(* IEC 61131-3 sources: PortalRobot/Portal_robot/Device/application/FB, 43 files *)

(* ---- F_GEOMETRY_EVENT.st ---- *)
FUNCTION F_GEOMETRY_EVENT : BOOL
VAR_INPUT
	Call : ST_GEOMETRY_CALL;
END_VAR
VAR
	uiIndex : UINT;
END_VAR

// --- BEGIN IMPLEMENTATION ---

// Один PLC-скан, единый владелец номера. Поля записываются раньше Seq.
Persistent_Value.udiEventSequence := Persistent_Value.udiEventSequence + UDINT#1;
IF Persistent_Value.udiEventSequence = UDINT#0 THEN Persistent_Value.udiEventSequence := UDINT#1; END_IF;
uiIndex := UDINT_TO_UINT((Persistent_Value.udiEventSequence - UDINT#1) MOD UDINT#100) + UINT#1;
GVL_GEOMETRY_CONTROL.astEvents[uiIndex].udiSequence := UDINT#0;
GVL_GEOMETRY_CONTROL.astEvents[uiIndex].Call := Call;
GVL_GEOMETRY_CONTROL.astEvents[uiIndex].udiTimeMs := GVL_HMI.udiHmiCommandClockMs;
GVL_GEOMETRY_CONTROL.astEvents[uiIndex].uiEnvironment := GVL_GEOMETRY_CONTROL.uiEnvironment;
GVL_GEOMETRY_CONTROL.astEvents[uiIndex].udiSequence := Persistent_Value.udiEventSequence;
F_GEOMETRY_EVENT := TRUE;

(* ---- F_GEOMETRY_SELECT_STATION.st ---- *)
FUNCTION F_GEOMETRY_SELECT_STATION : UINT
VAR_INPUT
	xRequireFree : BOOL;
	uiMachine : UINT := UINT#0; // Станок-источник; 0 — общая проверка доступности
END_VAR
VAR
	uiTry : UINT;
	uiStation : UINT;
END_VAR

// --- BEGIN IMPLEMENTATION ---

F_GEOMETRY_SELECT_STATION := UINT#0;
// С1/С2 предпочитают ГК1, С3 — ГК2. История доставок и магазины не участвуют.
uiStation := UINT#1;
IF uiMachine = UINT#3 THEN uiStation := UINT#2; END_IF;
FOR uiTry := UINT#1 TO UINT#2 DO
	// Вторым проверяем другой ГК, если предпочтительный не прошёл допуск.
	IF uiTry = UINT#2 THEN uiStation := UINT#3 - uiStation; END_IF;
	IF (F_GEOMETRY_SELECT_STATION = UINT#0) AND GVL_GEOMETRY_CONTROL.xSupported
	AND GVL_GEOMETRY_CONTROL.astStatus[uiStation].xEnabled
	AND NOT GVL_GEOMETRY_CONTROL.astStatus[uiStation].xDisablePending
	AND GVL_GEOMETRY_CONTROL.astStatus[uiStation].xConfigured
	AND NOT GVL_GEOMETRY_CONTROL.astStatus[uiStation].xError
	AND (GVL_GEOMETRY_CONTROL.astStatus[uiStation].uiState <> UINT#5) THEN
		IF NOT xRequireFree OR GVL_GEOMETRY_CONTROL.astStatus[uiStation].xReady THEN F_GEOMETRY_SELECT_STATION := uiStation; END_IF;
	END_IF;
END_FOR;

(* ---- F_GEOMETRY_TAKE_DETAIL.st ---- *)
FUNCTION F_GEOMETRY_TAKE_DETAIL : BOOL
VAR_INPUT
	uiMachine : UINT;
	uiProductType : UINT;
END_VAR
VAR
	Call : ST_GEOMETRY_CALL;
	EmptyCall : ST_GEOMETRY_CALL;
END_VAR

// --- BEGIN IMPLEMENTATION ---

F_GEOMETRY_TAKE_DETAIL := FALSE;
IF (uiMachine >= UINT#1) AND (uiMachine <= UINT#3) THEN
	// Считаем подтверждённую выгрузку ровно один раз, а не уровень Ready каждый скан.
	// Ожидающая выборка сохраняет счётчик до фактического взятия своей детали.
	IF (GVL_GEOMETRY_CONTROL.astCalls[uiMachine].uiState <> UINT#1)
	AND GVL_GEOMETRY_CONTROL.xSupported AND Persistent_Value.xAutoEnabled
	AND (GVL_GEOMETRY_CONTROL.astStatus[1].xEnabled OR GVL_GEOMETRY_CONTROL.astStatus[2].xEnabled) THEN
		GVL_GEOMETRY_CONTROL.auiActiveCount[uiMachine] := MIN(UINT#10000, GVL_GEOMETRY_CONTROL.auiActiveCount[uiMachine] + UINT#1);
		IF GVL_GEOMETRY_CONTROL.auiActiveCount[uiMachine] >= Persistent_Value.auiPeriod[uiMachine] THEN
			IF (GVL_GEOMETRY_CONTROL.astCalls[uiMachine].uiState <> UINT#2)
			AND (GVL_GEOMETRY_CONTROL.astCalls[uiMachine].uiState <> UINT#3) THEN
				Persistent_Value.udiNextCallId := Persistent_Value.udiNextCallId + UDINT#1;
				IF Persistent_Value.udiNextCallId = UDINT#0 THEN Persistent_Value.udiNextCallId := UDINT#1; END_IF;
				Call := EmptyCall; Call.udiId := Persistent_Value.udiNextCallId;
				Call.uiMachine := uiMachine; Call.uiProductType := uiProductType; Call.uiState := UINT#1;
				GVL_GEOMETRY_CONTROL.astCalls[uiMachine] := Call; F_GEOMETRY_EVENT(Call := Call);
			ELSE
				GVL_GEOMETRY_CONTROL.auiActiveCount[uiMachine] := UINT#0;
			END_IF;
		END_IF;
	END_IF;
	// Подхватываем вызов обслуживаемого станка независимо от вызовов других станков.
	// Повторная проверка после выезда также допускает поздний вызов своей детали.
	IF GVL_GEOMETRY_CONTROL.astCalls[uiMachine].uiState = UINT#1 THEN
		GVL_GEOMETRY_CONTROL.auiActiveCount[uiMachine] := UINT#0;
		GVL_GEOMETRY_CONTROL.astCalls[uiMachine].uiProductType := uiProductType;
		GVL_GEOMETRY_CONTROL.astCalls[uiMachine].uiState := UINT#2;
		F_GEOMETRY_EVENT(Call := GVL_GEOMETRY_CONTROL.astCalls[uiMachine]);
		F_GEOMETRY_TAKE_DETAIL := TRUE;
	END_IF;
END_IF;

(* ---- F_MAGAZINE_FRAME.st ---- *)
FUNCTION F_MAGAZINE_FRAME : ST_MAGAZINE_FRAME
VAR_INPUT
	stOrigin : ST_POINT;
	stCalibration : ST_MAGAZINE_CALIBRATION;
	uiRows : UINT;
	uiColumns : UINT;
	lrPitchX : LREAL;
	lrPitchY : LREAL;
END_VAR
VAR
	stFrame : ST_MAGAZINE_FRAME;
	stVectorAB : ST_MAGAZINE_VECTOR;
	stVectorAC : ST_MAGAZINE_VECTOR;
	stPlaneNormal : ST_MAGAZINE_VECTOR;
	lrVectorABLength : LREAL;
	lrPlaneNormalLength : LREAL;
END_VAR

// --- BEGIN IMPLEMENTATION ---

// Одноточечный режим сохраняет прежние направления мировых X/Y.
stFrame.stAxisX.X := 1.0; stFrame.stAxisX.Y := 0.0; stFrame.stAxisX.Z := 0.0;
stFrame.stAxisY.X := 0.0; stFrame.stAxisY.Y := 1.0; stFrame.stAxisY.Z := 0.0;
stFrame.stAxisZ.X := 0.0; stFrame.stAxisZ.Y := 0.0; stFrame.stAxisZ.Z := 1.0;
stFrame.xReady := FALSE;
stFrame.uiReason := UINT#0;
IF NOT stOrigin.xConfigured
OR (stOrigin.MagazineSafeZ = 0.0) OR (stOrigin.MagazineChangeZ = 0.0) THEN
	stFrame.uiReason := UINT#1;
ELSIF ((stCalibration.uiMethod <> UINT#1) AND (stCalibration.uiMethod <> UINT#3))
OR (uiRows = UINT#0) OR (uiColumns = UINT#0)
OR NOT ((lrPitchX >= 1.0) AND (lrPitchX <= 5000.0)
	AND (lrPitchY >= 1.0) AND (lrPitchY <= 5000.0)) THEN
	stFrame.uiReason := UINT#2;
ELSIF stCalibration.uiMethod = UINT#1 THEN
	stFrame.xReady := TRUE;
ELSIF (uiRows < UINT#2) OR (uiColumns < UINT#2) THEN
	stFrame.uiReason := UINT#2;
ELSIF NOT stCalibration.astReference[1].xConfigured
OR NOT stCalibration.astReference[2].xConfigured THEN
	stFrame.uiReason := UINT#3;
ELSE
	stVectorAB.X := stCalibration.astReference[1].X - stOrigin.X;
	stVectorAB.Y := stCalibration.astReference[1].Y - stOrigin.Y;
	stVectorAB.Z := stCalibration.astReference[1].Z - stOrigin.Z;
	stVectorAC.X := stCalibration.astReference[2].X - stOrigin.X;
	stVectorAC.Y := stCalibration.astReference[2].Y - stOrigin.Y;
	stVectorAC.Z := stCalibration.astReference[2].Z - stOrigin.Z;
	stPlaneNormal.X := stVectorAB.Y * stVectorAC.Z - stVectorAB.Z * stVectorAC.Y;
	stPlaneNormal.Y := stVectorAB.Z * stVectorAC.X - stVectorAB.X * stVectorAC.Z;
	stPlaneNormal.Z := stVectorAB.X * stVectorAC.Y - stVectorAB.Y * stVectorAC.X;
	lrVectorABLength := SQRT(stVectorAB.X * stVectorAB.X + stVectorAB.Y * stVectorAB.Y + stVectorAB.Z * stVectorAB.Z);
	lrPlaneNormalLength := SQRT(stPlaneNormal.X * stPlaneNormal.X + stPlaneNormal.Y * stPlaneNormal.Y + stPlaneNormal.Z * stPlaneNormal.Z);
	// Только математическая определённость: допуски размеров/углов не применяются.
	IF (lrVectorABLength > 0.0) AND (lrPlaneNormalLength > 0.0) THEN
		stFrame.stAxisX.X := stVectorAB.X / lrVectorABLength;
		stFrame.stAxisX.Y := stVectorAB.Y / lrVectorABLength;
		stFrame.stAxisX.Z := stVectorAB.Z / lrVectorABLength;
		stFrame.stAxisZ.X := stPlaneNormal.X / lrPlaneNormalLength;
		stFrame.stAxisZ.Y := stPlaneNormal.Y / lrPlaneNormalLength;
		stFrame.stAxisZ.Z := stPlaneNormal.Z / lrPlaneNormalLength;
		stFrame.stAxisY.X := stFrame.stAxisZ.Y * stFrame.stAxisX.Z - stFrame.stAxisZ.Z * stFrame.stAxisX.Y;
		stFrame.stAxisY.Y := stFrame.stAxisZ.Z * stFrame.stAxisX.X - stFrame.stAxisZ.X * stFrame.stAxisX.Z;
		stFrame.stAxisY.Z := stFrame.stAxisZ.X * stFrame.stAxisX.Y - stFrame.stAxisZ.Y * stFrame.stAxisX.X;
		// Сравнения также не принимают NaN/Inf после нечисловых входных данных.
		stFrame.xReady := (ABS(stFrame.stAxisX.X) <= 2.0) AND (ABS(stFrame.stAxisX.Y) <= 2.0)
			AND (ABS(stFrame.stAxisX.Z) <= 2.0) AND (ABS(stFrame.stAxisY.X) <= 2.0)
			AND (ABS(stFrame.stAxisY.Y) <= 2.0) AND (ABS(stFrame.stAxisY.Z) <= 2.0)
			AND (ABS(stFrame.stAxisZ.X) <= 2.0) AND (ABS(stFrame.stAxisZ.Y) <= 2.0)
			AND (ABS(stFrame.stAxisZ.Z) <= 2.0)
			AND ((stFrame.stAxisX.X * stFrame.stAxisX.X + stFrame.stAxisX.Y * stFrame.stAxisX.Y + stFrame.stAxisX.Z * stFrame.stAxisX.Z) > 0.0)
			AND ((stFrame.stAxisZ.X * stFrame.stAxisZ.X + stFrame.stAxisZ.Y * stFrame.stAxisZ.Y + stFrame.stAxisZ.Z * stFrame.stAxisZ.Z) > 0.0);
	END_IF;
	IF NOT stFrame.xReady THEN stFrame.uiReason := UINT#4; END_IF;
END_IF;
F_MAGAZINE_FRAME := stFrame;

(* ---- FB_ALARM_HORN.st ---- *)
FUNCTION_BLOCK FB_ALARM_HORN
VAR_INPUT
    astSource : ARRAY [1..22] OF ST_ALARM_SOURCE_DATA;
    tDuration : TIME := T#2S;
END_VAR
VAR_OUTPUT
    xSound : BOOL;
END_VAR
VAR
    adwPrevious : ARRAY [1..22] OF DWORD;
    uiSource : UINT;
    xNewAlarm : BOOL;
    xActive : BOOL;
    tLatchedDuration : TIME;
    tonSound : TON;
END_VAR

// --- BEGIN IMPLEMENTATION ---

// Предупреждения не входят в dwAlarmActive. Новая авария другого источника/бита
// тоже запускает звук, даже когда общая xAlarmActive уже была TRUE.
xNewAlarm := FALSE;
FOR uiSource := 1 TO 22 DO
    IF (astSource[uiSource].dwAlarmActive AND NOT adwPrevious[uiSource]) <> DWORD#0 THEN
        xNewAlarm := TRUE;
    END_IF;
    adwPrevious[uiSource] := astSource[uiSource].dwAlarmActive;
END_FOR;
IF tDuration <= T#0MS THEN
    xActive := FALSE;
ELSIF xNewAlarm THEN
    xActive := TRUE;
    tLatchedDuration := tDuration;
    // Сброс и запуск TON в этом же скане: новая авария начинает полный интервал.
    tonSound(IN := FALSE, PT := tLatchedDuration);
END_IF;
tonSound(IN := xActive, PT := tLatchedDuration);
IF tonSound.Q THEN
    xActive := FALSE;
END_IF;
xSound := xActive;

(* ---- FB_ALARM_MANAGER.st ---- *)
FUNCTION_BLOCK FB_ALARM_MANAGER
VAR_INPUT
	xResetWarnings : BOOL; // Сброс накопленных предупреждений
    xControllerWarningResetAllowed : BOOL; // 5C нельзя подтвердить до исчезновения свежей причины.
	astAdditionalCellWarning : ARRAY [1..2] OF ST_WARNING_EVENT; // Конфигуратор и ГК: независимые события источника CELL
END_VAR
VAR_IN_OUT
	Sources : ARRAY [1..22] OF ST_ALARM_SOURCE_DATA;
END_VAR
VAR_OUTPUT
    xEventsUpdated : BOOL; // Добавление, деактивация или подтверждение записи
	Status : ST_ALARM_STATUS; // Сводный статус журнала
	Events : ARRAY [1..100] OF ST_ALARM_EVENT; // Журнал активных и зафиксированных событий
END_VAR
VAR
    xSummaryInitialized : BOOL;
	uiWriteIndex : UINT := 1; // Следующая ячейка кольцевого журнала
	udiSequence  : UDINT; // Общий порядковый номер события
	adwPreviousAlarm : ARRAY [1..22] OF DWORD;
	audiPreviousWarning : ARRAY [1..22] OF UDINT;
	audiPreviousAdditionalCellWarning : ARRAY [1..2] OF UDINT;
	uiIndex : UINT; // Индекс источника или события
END_VAR

// --- BEGIN IMPLEMENTATION ---

xEventsUpdated := FALSE;

// Предупреждения подтверждаются только отдельной командой HMI.
// Общий сброс ошибок ячейки не изменяет журнал предупреждений.
IF xResetWarnings THEN
	FOR uiIndex := 1 TO 100 DO
		IF Events[uiIndex].xActive
		AND (Events[uiIndex].eSeverity = E_ALARM_SEVERITY.WARNING)
        AND ((Events[uiIndex].eSource <> E_ALARM_SOURCE.CONTROLLER_CPU_1)
            OR xControllerWarningResetAllowed) THEN
			Events[uiIndex].xActive := FALSE;
            xEventsUpdated := TRUE;
		END_IF;
	END_FOR;
END_IF;

// Менеджер не определяет причины: он регистрирует подготовленные данные владельцев блоков.
FOR uiIndex := 1 TO 22 DO
	UpdateSource(
		eSource := Sources[uiIndex].eSource,
		dwCurrent := Sources[uiIndex].dwAlarmActive,
		xRobotStopRequired := Sources[uiIndex].xRobotStopRequired,
		xGlobalError := Sources[uiIndex].xGlobalError,
		dwPrevious := adwPreviousAlarm[uiIndex]
	);

	IF Sources[uiIndex].stWarning.udiSequence <> audiPreviousWarning[uiIndex] THEN
		IF (Sources[uiIndex].stWarning.udiSequence <> UDINT#0)
		AND (Sources[uiIndex].stWarning.uiCode <> UINT#0) THEN
		AddEvent(
			eSource := Sources[uiIndex].eSource,
			eSeverity := E_ALARM_SEVERITY.WARNING,
			eEffect := E_ALARM_EFFECT.WARNING,
			uiCode := Sources[uiIndex].stWarning.uiCode
		);
		END_IF;
		audiPreviousWarning[uiIndex] := Sources[uiIndex].stWarning.udiSequence;
	END_IF;
END_FOR;

// Общие предупреждения ГК и конфигуратора не изменяют последний код/счётчик
// FB_CELL_MANAGER. Иначе возврат его старого снимка становился новым событием.
// Обрабатываем все каналы в одном вызове: события одного скана не теряются,
// а xResetWarnings не очищает предупреждение, выданное после сброса в этом скане.
FOR uiIndex := UINT#1 TO UINT#2 DO
	IF astAdditionalCellWarning[uiIndex].udiSequence <> audiPreviousAdditionalCellWarning[uiIndex] THEN
		IF (astAdditionalCellWarning[uiIndex].udiSequence <> UDINT#0)
		AND (astAdditionalCellWarning[uiIndex].uiCode <> UINT#0) THEN
			AddEvent(
				eSource := E_ALARM_SOURCE.CELL,
				eSeverity := E_ALARM_SEVERITY.WARNING,
				eEffect := E_ALARM_EFFECT.WARNING,
				uiCode := astAdditionalCellWarning[uiIndex].uiCode
			);
		END_IF;
		audiPreviousAdditionalCellWarning[uiIndex] := astAdditionalCellWarning[uiIndex].udiSequence;
	END_IF;
END_FOR;

IF xEventsUpdated OR NOT xSummaryInitialized THEN
Status.uiActiveAlarmCount := 0;
Status.uiActiveWarningCount := 0;
Status.uiHistoryCount := 0;

FOR uiIndex := 1 TO 100 DO
	IF Events[uiIndex].udiSequence <> UDINT#0 THEN
		Status.uiHistoryCount := Status.uiHistoryCount + 1;
	END_IF;
	IF Events[uiIndex].xActive THEN
		IF Events[uiIndex].eSeverity = E_ALARM_SEVERITY.ALARM THEN
			Status.uiActiveAlarmCount := Status.uiActiveAlarmCount + 1;
		ELSE
			Status.uiActiveWarningCount := Status.uiActiveWarningCount + 1;
		END_IF;
	END_IF;
END_FOR;

Status.uiActiveEventCount := Status.uiActiveAlarmCount + Status.uiActiveWarningCount;
Status.xAlarmActive := Status.uiActiveAlarmCount > 0;
Status.xWarningActive := Status.uiActiveWarningCount > 0;
    xSummaryInitialized := TRUE;
END_IF;

(* ---- FB_AXIS.st ---- *)
FUNCTION_BLOCK FB_Axis
VAR_INPUT
	FaultRequest : ST_AXIS_FAULT_REQUEST; // Единый контракт диагностической инъекции
	xResetPermit : BOOL; // Общий сброс разрешён ручным режимом и остановленной ячейкой
END_VAR
VAR_OUTPUT
	FaultStatus : ST_FAULT_INJECTION_STATUS; // Состояние инжектора для HMI
END_VAR
VAR_IN_OUT
    Axis     : AXIS_REF_SM3;   // ссылка на ось SoftMotion
    AxisData : ST_AXIS;        // все данные оси (команды, параметры, статусы)
END_VAR

VAR CONSTANT
    // ==================================================
    // Ошибки оси, MC-блоков и SoftMotion
    // ==================================================
    AXE_MC_POWER_ERROR       : DWORD := DWORD#16#00000001; // Ошибка MC_Power
    AXE_MC_RESET_ERROR       : DWORD := DWORD#16#00000002; // Ошибка MC_Reset
    AXE_MC_STOP_ERROR        : DWORD := DWORD#16#00000004; // Ошибка MC_Stop
    AXE_MC_JOG_ERROR         : DWORD := DWORD#16#00000008; // Ошибка MC_Jog
    AXE_MC_HOME_ERROR        : DWORD := DWORD#16#00000010; // Ошибка MC_Home
    AXE_MC_MOVE_ABS_ERROR    : DWORD := DWORD#16#00000020; // Ошибка абсолютного перемещения
    AXE_MC_MOVE_REL_ERROR    : DWORD := DWORD#16#00000040; // Ошибка относительного перемещения
    AXE_READ_POS_ERROR       : DWORD := DWORD#16#00000080; // Ошибка чтения позиции
    AXE_READ_STATUS_ERROR    : DWORD := DWORD#16#00000100; // Ошибка чтения статуса
    AXE_ERRORSTOP            : DWORD := DWORD#16#00000200; // Ось находится в ErrorStop
    AXE_FB_ERROR_OCCURRED    : DWORD := DWORD#16#00000400; // SoftMotion сообщил внутреннюю ошибку
    AXE_COMMAND_ABORTED      : DWORD := DWORD#16#00000800; // Команда движения прервана
    AXE_UNKNOWN_ACTUAL_ERROR : DWORD := DWORD#16#00001000; // Неизвестная текущая ошибка
    AXE_DRIVE_AXIS_ERROR     : DWORD := DWORD#16#00002000; // Ошибка привода
    AXE_POWER_FEEDBACK_LOST  : DWORD := DWORD#16#00004000; // Потеря силовой готовности при активной команде питания

    // ==================================================
    // Логические ошибки блока
    // ==================================================
    LOG_POWER_PERMIT_LOST    : DWORD := DWORD#16#00000001; // Снято разрешение питания
    LOG_GLOBAL_DURING_POWER  : DWORD := DWORD#16#00000002; // Глобальная ошибка при включении
    LOG_GLOBAL_DURING_READY  : DWORD := DWORD#16#00000004; // Глобальная ошибка в готовности
    LOG_GLOBAL_DURING_MOTION : DWORD := DWORD#16#00000008; // Глобальная ошибка при движении
    LOG_JOG_CONFLICT         : DWORD := DWORD#16#00000010; // Одновременно заданы Jog+ и Jog-
    LOG_MOVE_ABS_NOT_HOMED   : DWORD := DWORD#16#00000020; // Абсолютное движение без поиска дома
    LOG_MOVE_REL_NOT_HOMED   : DWORD := DWORD#16#00000040; // Относительное движение без поиска дома
    LOG_STEP_TIMEOUT         : DWORD := DWORD#16#00000080; // Превышено время шага
    LOG_UNKNOWN_STEP         : DWORD := DWORD#16#00000100; // Неизвестный шаг автомата

    // ==================================================
    // Предупреждения блока
    // ==================================================
    WRN_NO_POWER_PERMIT : DWORD := DWORD#16#00000001; // Нет разрешения подачи питания
    WRN_RESET_GLOBAL_ERROR   : UINT := 2; // Сброс не выполнен из-за глобальной ошибки
    WRN_RESET_MC_ERROR       : UINT := 3; // MC_Reset завершился ошибкой
    WRN_RESET_TIMEOUT        : UINT := 4; // Превышено время сброса
    WRN_RESET_AXIS_ACTIVE    : UINT := 5; // Физическая ошибка оси осталась активной
    WRN_RESET_AXIS_LATCHED   : UINT := 6; // Защёлкнутая ошибка оси не была очищена
    WRN_RESET_LOGICAL_ACTIVE : UINT := 7; // Логическая ошибка оси не была очищена
	WRN_SIM_ERROR_NOT_ALLOWED : UINT := 8; // Тестовый конфликт Jog запрещён состоянием оси

END_VAR

VAR
	lrEffectiveVelocity : LREAL;
	lrEffectiveAcceleration : LREAL;
	lrEffectiveDeceleration : LREAL;
	lrEffectiveJerk : LREAL;
    // Триггеры на команды
    rtEnable            : R_TRIG; // Фронт команды включения
    rtDisable           : R_TRIG; // Фронт команды отключения
    rtResetAllError     : R_TRIG; // Фронт общего сброса
    rtResetAxisError    : R_TRIG; // Фронт сброса привода
    rtResetLogicalError : R_TRIG; // Фронт сброса логики
    rtStop              : R_TRIG; // Фронт команды остановки
    rtHome              : R_TRIG; // Фронт команды поиска дома
    rtMoveAbsolute      : R_TRIG; // Фронт абсолютного перемещения
    rtMoveRelative      : R_TRIG; // Фронт относительного перемещения

    // Экземпляры MC-блоков
    fbPower        : MC_Power; // Управление питанием привода
    fbReset        : MC_Reset; // Сброс ошибки привода
    fbStop         : MC_Stop; // Контролируемая остановка
    fbJog          : MC_Jog; // Толчковое движение
    fbHome         : MC_Home; // Поиск домашней позиции
    fbMoveAbsolute : MC_MoveAbsolute; // Абсолютное перемещение
    fbMoveRelative : MC_MoveRelative; // Относительное перемещение
    fbReadPosition : MC_ReadActualPosition; // Чтение текущей позиции
    fbReadStatus   : MC_ReadStatus; // Чтение состояния оси
    fbReadAxisError: MC_ReadAxisError; // Чтение кода ошибки привода

    // Внутренние управляющие флаги
    xPowerRequest    : BOOL; // Защёлкнутый запрос питания
    xResetExecute    : BOOL; // Выполняется сброс привода
    xStopExecute     : BOOL; // Выполняется остановка
    xHomeExecute     : BOOL; // Выполняется поиск дома
    xMoveAbsExecute  : BOOL; // Выполняется абсолютное перемещение
    xMoveRelExecute  : BOOL; // Выполняется относительное перемещение
    xJogForwardExec  : BOOL; // Выполняется Jog в положительную сторону
    xJogBackwardExec : BOOL; // Выполняется Jog в отрицательную сторону

    // Для таймера шага
    iPrevStep        : E_AXIS_STATE := E_AXIS_STATE.DISABLED; // Предыдущий шаг автомата
    xStepChanged     : BOOL; // Шаг изменился в текущем цикле
    xStepTimerEnable : BOOL; // Разрешение таймера шага
    tonStep          : TON; // Таймер времени на шаге
    tonStepTimeout   : TON; // Таймер превышения времени шага
    tonPowerFeedbackLoss : TON; // Контроль неожиданного снятия силовой готовности
    xPowerFeedbackExpected : BOOL; // Текущее состояние требует сохранения питания

    // Для удержания предупреждений
    tpWarningHold : TP; // Удержание предупреждения для отображения
    xWarningPulse : BOOL; // Импульс нового предупреждения

    // Вспомогательные флаги для сброса
    xDoResetAxis    : BOOL; // Требуется сброс ошибок привода
    xDoResetLogical : BOOL; // Требуется сброс логических ошибок
    xNeedMcReset    : BOOL; // Требуется вызов MC_Reset
    uiResetWarningCode : UINT; // Причина неуспешного сброса текущего цикла

    // Актуальная ошибка оси (на основе MC-блоков)
    xAxisErrorActual : BOOL; // Текущая ошибка по выходам MC-блоков
	fbFaultInjector : FB_AXIS_FAULT_INJECTOR; // Безопасный источник логической ошибки Jog
	xFaultAllowed   : BOOL; // Условия теста, рассчитанные владельцем оси
END_VAR

// --- BEGIN IMPLEMENTATION ---

// Коэффициент симуляции не изменяет динамику осей робота.
// Скорость, ускорение, замедление и jerk задаются пользователем в настройках осей.
lrEffectiveVelocity := AxisData.MotionParam.lrVelocity;
lrEffectiveAcceleration := AxisData.MotionParam.lrAcceleration;
lrEffectiveDeceleration := AxisData.MotionParam.lrDeceleration;
lrEffectiveJerk := AxisData.MotionParam.lrJerk;

// ======================================================
// 1. ФРОНТЫ (триггеры на команды из структуры)
// ======================================================
rtEnable(CLK := AxisData.Command.xEnable);
rtDisable(CLK := AxisData.Command.xDisable);
rtResetAllError(CLK := AxisData.Command.xResetAllError);
rtResetAxisError(CLK := AxisData.Command.xResetAxisError);
rtResetLogicalError(CLK := AxisData.Command.xResetLogicalError);
rtStop(CLK := AxisData.Command.xStop);
rtHome(CLK := AxisData.Command.xHome);
rtMoveAbsolute(CLK := AxisData.Command.xMoveAbsolute);
rtMoveRelative(CLK := AxisData.Command.xMoveRelative);

// ======================================================
// 2. СТАТУСЫ ОТ MC-БЛОКОВ (запись в структуру)
// ======================================================
AxisData.Status.xPowerStageOn := fbPower.bRegulatorRealState;
AxisData.Status.xDriveStartOn := fbPower.bDriveStartRealState;
AxisData.Status.xPowered := fbPower.Status
	AND AxisData.Status.xPowerStageOn
	AND AxisData.Status.xDriveStartOn;
AxisData.Status.xPowerOff := NOT AxisData.Status.xPowerStageOn
	AND NOT AxisData.Status.xDriveStartOn;

AxisData.Status.xLocalError :=
    fbPower.Error OR
    fbReset.Error OR
    fbStop.Error OR
    fbJog.Error OR
    fbHome.Error OR
    fbMoveAbsolute.Error OR
    fbMoveRelative.Error OR
    fbReadPosition.Error OR
    fbReadStatus.Error OR
    fbReadStatus.Errorstop OR
    fbReadStatus.FBErrorOccured;

AxisData.Status.xMotionBusy :=
    fbStop.Busy OR
    fbJog.Busy OR
    fbHome.Busy OR
    fbMoveAbsolute.Busy OR
    fbMoveRelative.Busy;

// MC_Reset нужен только для аппаратных/SoftMotion ошибок
xNeedMcReset := fbReadStatus.Errorstop OR fbReadStatus.FBErrorOccured OR fbReadAxisError.AxisError;

AxisData.Error.dwAxisError := AxisData.Error.dwAxisErrorActual OR AxisData.Error.dwAxisErrorLatched;
AxisData.Error.dwLogicalError := AxisData.Error.dwLogicalErrorLatched;
AxisData.Error.dwAllError := AxisData.Error.dwAxisError OR AxisData.Error.dwLogicalError;

// ======================================================
// 3. ЗНАЧЕНИЯ ПО УМОЛЧАНИЮ ДЛЯ ИСПОЛНИТЕЛЬНЫХ ФЛАГОВ
// ======================================================
xResetExecute    := FALSE;
xStopExecute     := FALSE;
xHomeExecute     := FALSE;
xMoveAbsExecute  := FALSE;
xMoveRelExecute  := FALSE;
xJogForwardExec  := FALSE;
xJogBackwardExec := FALSE;

AxisData.Status.xDone := FALSE;
xWarningPulse := FALSE;
uiResetWarningCode := UINT#0;

// MC_Power не обязан выставлять Error при отказе интерфейса привода. Например,
// окончание demo-лицензии SoftMotion снимает реальные Regulator/DriveStart,
// но оставляет AxisError и FBError пустыми. Контролируем поэтому сам факт
// исчезновения силовой готовности при сохраняющемся запросе питания.
xPowerFeedbackExpected := xPowerRequest
	AND AxisData.Command.xPowerPermit
	AND ((AxisData.Diag.iStep = E_AXIS_STATE.READY)
		OR (AxisData.Diag.iStep = E_AXIS_STATE.JOGGING)
		OR (AxisData.Diag.iStep = E_AXIS_STATE.JOG_DECELERATING)
		OR (AxisData.Diag.iStep = E_AXIS_STATE.HOMING)
		OR (AxisData.Diag.iStep = E_AXIS_STATE.MOVE_ABSOLUTE)
		OR (AxisData.Diag.iStep = E_AXIS_STATE.MOVE_RELATIVE)
		OR (AxisData.Diag.iStep = E_AXIS_STATE.STOPPING)
		OR (AxisData.Diag.iStep = E_AXIS_STATE.STOP_RELEASE));
tonPowerFeedbackLoss(
	IN := xPowerFeedbackExpected AND NOT AxisData.Status.xPowered,
	PT := AxisData.Timeouts.tPowerFeedbackLossTimeout
);
IF tonPowerFeedbackLoss.Q
AND (AxisData.Diag.iStep <> E_AXIS_STATE.ERROR_RESET_MANAGER) THEN
	AxisData.Error.dwAxisErrorLatched :=
		AxisData.Error.dwAxisErrorLatched OR AXE_POWER_FEEDBACK_LOST;
	AxisData.Diag.iLastErrorStep := TO_INT(AxisData.Diag.iStep);
	AxisData.Diag.iStep := E_AXIS_STATE.ERROR_RESET_MANAGER;
END_IF;

// Конфликт Jog проверяется автоматом до вызова MC_Jog, поэтому тест не создаёт движения.
xFaultAllowed := (AxisData.Diag.iStep = E_AXIS_STATE.READY)
	AND NOT AxisData.Command.xGlobalError
	AND NOT AxisData.Status.xError
	AND NOT AxisData.Status.xMotionBusy
	AND NOT AxisData.Command.xJogPositive
	AND NOT AxisData.Command.xJogNegative
	AND NOT AxisData.Command.xHome
	AND NOT AxisData.Command.xMoveAbsolute
	AND NOT AxisData.Command.xMoveRelative;

fbFaultInjector(
	Request := FaultRequest,
	xOwnerAllowed := xFaultAllowed
);
FaultStatus := fbFaultInjector.Status;

IF fbFaultInjector.Status.xRejected THEN
	AxisData.Diag.sWarningText := 'Simulated Jog conflict is not allowed';
	AxisData.Diag.stWarning.uiCode := WRN_SIM_ERROR_NOT_ALLOWED;
	AxisData.Diag.stWarning.udiSequence := AxisData.Diag.stWarning.udiSequence + UDINT#1;
	IF AxisData.Diag.stWarning.udiSequence = UDINT#0 THEN
		AxisData.Diag.stWarning.udiSequence := UDINT#1;
	END_IF;
	xWarningPulse := TRUE;
END_IF;

// ======================================================
// 4. КОНЕЧНЫЙ АВТОМАТ (используем перечисление E_AXIS_STATE)
// ======================================================
CASE AxisData.Diag.iStep OF

    // --------------------------------------------------
    E_AXIS_STATE.DISABLED:
    // --------------------------------------------------
        AxisData.Diag.sStepName := 'DISABLED';
        AxisData.Diag.sWaitReason := 'Waiting Enable command';
        AxisData.Diag.tStepPreset := T#0S;

        xPowerRequest := FALSE;
        AxisData.Status.xHomed := FALSE;

        IF AxisData.Status.xError THEN
            AxisData.Diag.iStep := E_AXIS_STATE.ERROR_RESET_MANAGER;

        ELSIF rtEnable.Q AND NOT AxisData.Command.xPowerPermit THEN
            AxisData.Error.dwWarningLatched :=
                AxisData.Error.dwWarningLatched OR WRN_NO_POWER_PERMIT;
            AxisData.Diag.sWarningText := 'Power permit is not active';
            AxisData.Diag.stWarning.uiCode := UINT#1;
            AxisData.Diag.stWarning.udiSequence := AxisData.Diag.stWarning.udiSequence + UDINT#1;
            IF AxisData.Diag.stWarning.udiSequence = UDINT#0 THEN
                AxisData.Diag.stWarning.udiSequence := UDINT#1;
            END_IF;
            xWarningPulse := TRUE;
            AxisData.Diag.sWaitReason := 'Power permit missing';

        ELSIF NOT AxisData.Command.xPowerPermit THEN
            AxisData.Diag.sWaitReason := 'Power permit missing';

        ELSIF rtEnable.Q THEN
            xPowerRequest := TRUE;
            AxisData.Diag.iStep := E_AXIS_STATE.POWERING;
        END_IF;

    // --------------------------------------------------
    E_AXIS_STATE.POWERING:
    // --------------------------------------------------
        AxisData.Diag.sStepName := 'POWERING';
        AxisData.Diag.sWaitReason := 'Waiting MC_Power.Status';
        AxisData.Diag.tStepPreset := AxisData.Timeouts.tPowerTimeout;

        xPowerRequest := TRUE;

        IF NOT AxisData.Command.xPowerPermit THEN
            xPowerRequest := FALSE;
            AxisData.Error.dwLogicalErrorLatched :=
                AxisData.Error.dwLogicalErrorLatched OR LOG_POWER_PERMIT_LOST;
            AxisData.Diag.iLastErrorStep := TO_INT(AxisData.Diag.iStep);
            AxisData.Diag.iStep := E_AXIS_STATE.ERROR_RESET_MANAGER;

        ELSIF AxisData.Command.xGlobalError THEN
            xPowerRequest := FALSE;
            AxisData.Error.dwLogicalErrorLatched :=
                AxisData.Error.dwLogicalErrorLatched OR LOG_GLOBAL_DURING_POWER;
            AxisData.Diag.iLastErrorStep := TO_INT(AxisData.Diag.iStep);
            AxisData.Diag.iStep := E_AXIS_STATE.ERROR_RESET_MANAGER;

        ELSIF fbPower.Error THEN
            xPowerRequest := FALSE;
            AxisData.Error.dwAxisErrorLatched :=
                AxisData.Error.dwAxisErrorLatched OR AXE_MC_POWER_ERROR;
            AxisData.Diag.udiLastErrorID := TO_UDINT(fbPower.ErrorID);
            AxisData.Diag.iLastErrorStep := TO_INT(AxisData.Diag.iStep);
            AxisData.Diag.iStep := E_AXIS_STATE.ERROR_RESET_MANAGER;

        // READY допустим только после подтверждения всех трёх признаков:
        // MC_Power.Status, силовая ступень и снятый quickstop.
        ELSIF AxisData.Status.xPowered THEN
            AxisData.Diag.iStep := E_AXIS_STATE.READY;

        ELSIF rtDisable.Q THEN
            xPowerRequest := FALSE;
            AxisData.Diag.iStep := E_AXIS_STATE.POWERING_DOWN;
        END_IF;

    // --------------------------------------------------
    E_AXIS_STATE.POWERING_DOWN:
    // --------------------------------------------------
        AxisData.Diag.sStepName := 'POWERING_DOWN';
        AxisData.Diag.sWaitReason := 'Waiting drive power feedback off';
        AxisData.Diag.tStepPreset := AxisData.Timeouts.tPowerTimeout;

        xPowerRequest := FALSE;

        IF fbPower.Error THEN
            AxisData.Error.dwAxisErrorLatched :=
                AxisData.Error.dwAxisErrorLatched OR AXE_MC_POWER_ERROR;
            AxisData.Diag.udiLastErrorID := TO_UDINT(fbPower.ErrorID);
            AxisData.Diag.iLastErrorStep := TO_INT(AxisData.Diag.iStep);
            AxisData.Diag.iStep := E_AXIS_STATE.ERROR_RESET_MANAGER;

        ELSIF AxisData.Status.xPowerOff THEN
            AxisData.Diag.iStep := E_AXIS_STATE.DISABLED;
        END_IF;

    // --------------------------------------------------
    E_AXIS_STATE.READY:
    // --------------------------------------------------
        AxisData.Diag.sStepName := 'READY';
        AxisData.Diag.sWaitReason := 'Waiting command';
        AxisData.Diag.tStepPreset := T#0S;

        xPowerRequest := TRUE;

        IF NOT AxisData.Command.xPowerPermit THEN
            xPowerRequest := FALSE;
            AxisData.Diag.iStep := E_AXIS_STATE.POWERING_DOWN;

        ELSIF rtDisable.Q THEN
            xPowerRequest := FALSE;
            AxisData.Diag.iStep := E_AXIS_STATE.POWERING_DOWN;

        ELSIF AxisData.Command.xGlobalError THEN
            AxisData.Error.dwLogicalErrorLatched :=
                AxisData.Error.dwLogicalErrorLatched OR LOG_GLOBAL_DURING_READY;
            AxisData.Diag.iLastErrorStep := TO_INT(AxisData.Diag.iStep);
            AxisData.Diag.iStep := E_AXIS_STATE.ERROR_RESET_MANAGER;

        ELSIF xAxisErrorActual THEN
            AxisData.Error.dwAxisErrorLatched :=
                AxisData.Error.dwAxisErrorLatched OR AxisData.Error.dwAxisErrorActual;
            AxisData.Diag.iLastErrorStep := TO_INT(AxisData.Diag.iStep);
            AxisData.Diag.iStep := E_AXIS_STATE.ERROR_RESET_MANAGER;

        ELSIF fbFaultInjector.xJogConflict
		OR (AxisData.Command.xJogPositive AND AxisData.Command.xJogNegative) THEN
            AxisData.Error.dwLogicalErrorLatched :=
                AxisData.Error.dwLogicalErrorLatched OR LOG_JOG_CONFLICT;
            AxisData.Diag.iLastErrorStep := TO_INT(AxisData.Diag.iStep);
            AxisData.Diag.iStep := E_AXIS_STATE.ERROR_RESET_MANAGER;

        ELSIF AxisData.Command.xJogPositive OR AxisData.Command.xJogNegative THEN
            AxisData.Diag.iStep := E_AXIS_STATE.JOGGING;

        ELSIF rtHome.Q THEN
            AxisData.Diag.iStep := E_AXIS_STATE.HOMING;

        ELSIF rtMoveAbsolute.Q THEN
            IF AxisData.Status.xHomed THEN
                AxisData.Diag.iStep := E_AXIS_STATE.MOVE_ABSOLUTE;
            ELSE
                AxisData.Error.dwLogicalErrorLatched :=
                    AxisData.Error.dwLogicalErrorLatched OR LOG_MOVE_ABS_NOT_HOMED;
                AxisData.Diag.iLastErrorStep := TO_INT(AxisData.Diag.iStep);
                AxisData.Diag.iStep := E_AXIS_STATE.ERROR_RESET_MANAGER;
            END_IF;

        ELSIF rtMoveRelative.Q THEN
            IF AxisData.Status.xHomed THEN
                AxisData.Diag.iStep := E_AXIS_STATE.MOVE_RELATIVE;
            ELSE
                AxisData.Error.dwLogicalErrorLatched :=
                    AxisData.Error.dwLogicalErrorLatched OR LOG_MOVE_REL_NOT_HOMED;
                AxisData.Diag.iLastErrorStep := TO_INT(AxisData.Diag.iStep);
                AxisData.Diag.iStep := E_AXIS_STATE.ERROR_RESET_MANAGER;
            END_IF;
        END_IF;

    // --------------------------------------------------
    E_AXIS_STATE.JOGGING:
    // --------------------------------------------------
        AxisData.Diag.sStepName := 'JOGGING';
        AxisData.Diag.sWaitReason := 'Jog active';
        AxisData.Diag.tStepPreset := T#0S;

        xPowerRequest := TRUE;
        xJogForwardExec  := AxisData.Command.xJogPositive AND NOT AxisData.Command.xJogNegative;
        xJogBackwardExec := AxisData.Command.xJogNegative AND NOT AxisData.Command.xJogPositive;

        IF NOT AxisData.Command.xPowerPermit THEN
            xJogForwardExec := FALSE;
            xJogBackwardExec := FALSE;
            AxisData.Error.dwLogicalErrorLatched :=
                AxisData.Error.dwLogicalErrorLatched OR LOG_POWER_PERMIT_LOST;
            AxisData.Diag.iLastErrorStep := TO_INT(AxisData.Diag.iStep);
            AxisData.Diag.iStep := E_AXIS_STATE.STOPPING;

        ELSIF AxisData.Command.xGlobalError THEN
            xJogForwardExec := FALSE;
            xJogBackwardExec := FALSE;
            AxisData.Error.dwLogicalErrorLatched :=
                AxisData.Error.dwLogicalErrorLatched OR LOG_GLOBAL_DURING_MOTION;
            AxisData.Diag.iLastErrorStep := TO_INT(AxisData.Diag.iStep);
            AxisData.Diag.iStep := E_AXIS_STATE.STOPPING;

        ELSIF xAxisErrorActual THEN
            xJogForwardExec := FALSE;
            xJogBackwardExec := FALSE;
            AxisData.Error.dwAxisErrorLatched :=
                AxisData.Error.dwAxisErrorLatched OR AxisData.Error.dwAxisErrorActual;
            AxisData.Diag.iLastErrorStep := TO_INT(AxisData.Diag.iStep);
            // SoftMotion уже перевёл ось в ErrorStop и выполнил error ramp.
            // MC_Stop в этом состоянии создаёт вторичную ошибку "axis is in errorstop".
            AxisData.Diag.iStep := E_AXIS_STATE.ERROR_RESET_MANAGER;

        ELSIF rtStop.Q THEN
            xJogForwardExec := FALSE;
            xJogBackwardExec := FALSE;
            AxisData.Diag.iStep := E_AXIS_STATE.STOPPING;

        ELSIF AxisData.Command.xJogPositive AND AxisData.Command.xJogNegative THEN
            xJogForwardExec := FALSE;
            xJogBackwardExec := FALSE;
            AxisData.Error.dwLogicalErrorLatched :=
                AxisData.Error.dwLogicalErrorLatched OR LOG_JOG_CONFLICT;
            AxisData.Diag.iLastErrorStep := TO_INT(AxisData.Diag.iStep);
            AxisData.Diag.iStep := E_AXIS_STATE.STOPPING;

        ELSIF NOT AxisData.Command.xJogPositive AND NOT AxisData.Command.xJogNegative THEN
            xJogForwardExec := FALSE;
            xJogBackwardExec := FALSE;
            AxisData.Diag.iStep := E_AXIS_STATE.JOG_DECELERATING;
        END_IF;

    // --------------------------------------------------
    E_AXIS_STATE.JOG_DECELERATING:
    // --------------------------------------------------
        AxisData.Diag.sStepName := 'JOG_DECELERATING';
        AxisData.Diag.sWaitReason := 'Waiting MC_Jog controlled deceleration';
        AxisData.Diag.tStepPreset := T#0S;

        xPowerRequest := TRUE;
        xJogForwardExec := FALSE;
        xJogBackwardExec := FALSE;

        IF NOT AxisData.Command.xPowerPermit THEN
            AxisData.Error.dwLogicalErrorLatched :=
                AxisData.Error.dwLogicalErrorLatched OR LOG_POWER_PERMIT_LOST;
            AxisData.Diag.iLastErrorStep := TO_INT(AxisData.Diag.iStep);
            AxisData.Diag.iStep := E_AXIS_STATE.STOPPING;

        ELSIF AxisData.Command.xGlobalError THEN
            AxisData.Error.dwLogicalErrorLatched :=
                AxisData.Error.dwLogicalErrorLatched OR LOG_GLOBAL_DURING_MOTION;
            AxisData.Diag.iLastErrorStep := TO_INT(AxisData.Diag.iStep);
            AxisData.Diag.iStep := E_AXIS_STATE.STOPPING;

        ELSIF xAxisErrorActual THEN
            AxisData.Error.dwAxisErrorLatched :=
                AxisData.Error.dwAxisErrorLatched OR AxisData.Error.dwAxisErrorActual;
            AxisData.Diag.iLastErrorStep := TO_INT(AxisData.Diag.iStep);
            AxisData.Diag.iStep := E_AXIS_STATE.ERROR_RESET_MANAGER;

        ELSIF rtStop.Q THEN
            AxisData.Diag.iStep := E_AXIS_STATE.STOPPING;

        ELSIF AxisData.Command.xJogPositive AND AxisData.Command.xJogNegative THEN
            AxisData.Error.dwLogicalErrorLatched :=
                AxisData.Error.dwLogicalErrorLatched OR LOG_JOG_CONFLICT;
            AxisData.Diag.iLastErrorStep := TO_INT(AxisData.Diag.iStep);
            AxisData.Diag.iStep := E_AXIS_STATE.STOPPING;

        ELSIF AxisData.Command.xJogPositive OR AxisData.Command.xJogNegative THEN
            AxisData.Diag.iStep := E_AXIS_STATE.JOGGING;

        ELSIF NOT fbJog.Busy THEN
            AxisData.Status.xDone := TRUE;
            AxisData.Diag.iStep := E_AXIS_STATE.READY;
        END_IF;

    // --------------------------------------------------
    E_AXIS_STATE.HOMING:
    // --------------------------------------------------
        AxisData.Diag.sStepName := 'HOMING';
        AxisData.Diag.sWaitReason := 'Waiting MC_Home.Done';
        AxisData.Diag.tStepPreset := AxisData.Timeouts.tHomeTimeout;

        xPowerRequest := TRUE;
        xHomeExecute := TRUE;

        IF NOT AxisData.Command.xPowerPermit THEN
            xHomeExecute := FALSE;
            AxisData.Error.dwLogicalErrorLatched :=
                AxisData.Error.dwLogicalErrorLatched OR LOG_POWER_PERMIT_LOST;
            AxisData.Diag.iLastErrorStep := TO_INT(AxisData.Diag.iStep);
            AxisData.Diag.iStep := E_AXIS_STATE.STOPPING;

        ELSIF AxisData.Command.xGlobalError THEN
            xHomeExecute := FALSE;
            AxisData.Error.dwLogicalErrorLatched :=
                AxisData.Error.dwLogicalErrorLatched OR LOG_GLOBAL_DURING_MOTION;
            AxisData.Diag.iLastErrorStep := TO_INT(AxisData.Diag.iStep);
            AxisData.Diag.iStep := E_AXIS_STATE.STOPPING;

        ELSIF rtStop.Q THEN
            xHomeExecute := FALSE;
            AxisData.Diag.iStep := E_AXIS_STATE.STOPPING;

        ELSIF fbHome.Error THEN
            xHomeExecute := FALSE;
            AxisData.Error.dwAxisErrorLatched :=
                AxisData.Error.dwAxisErrorLatched OR AXE_MC_HOME_ERROR;
            AxisData.Diag.udiLastErrorID := TO_UDINT(fbHome.ErrorID);
            AxisData.Diag.iLastErrorStep := TO_INT(AxisData.Diag.iStep);
            AxisData.Diag.iStep := E_AXIS_STATE.ERROR_RESET_MANAGER;

        ELSIF fbHome.CommandAborted THEN
            xHomeExecute := FALSE;
            AxisData.Error.dwAxisErrorLatched :=
                AxisData.Error.dwAxisErrorLatched OR AXE_COMMAND_ABORTED;
            AxisData.Diag.udiLastErrorID := 3003;
            AxisData.Diag.iLastErrorStep := TO_INT(AxisData.Diag.iStep);
            AxisData.Diag.iStep := E_AXIS_STATE.ERROR_RESET_MANAGER;

        ELSIF xAxisErrorActual THEN
            xHomeExecute := FALSE;
            AxisData.Error.dwAxisErrorLatched :=
                AxisData.Error.dwAxisErrorLatched OR AxisData.Error.dwAxisErrorActual;
            AxisData.Diag.iLastErrorStep := TO_INT(AxisData.Diag.iStep);
            AxisData.Diag.iStep := E_AXIS_STATE.ERROR_RESET_MANAGER;

        ELSIF fbHome.Done THEN
            xHomeExecute := FALSE;
            AxisData.Status.xHomed := TRUE;
            AxisData.Status.xDone := TRUE;
            AxisData.Diag.iStep := E_AXIS_STATE.READY;
        END_IF;

    // --------------------------------------------------
    E_AXIS_STATE.MOVE_ABSOLUTE:
    // --------------------------------------------------
        AxisData.Diag.sStepName := 'MOVING_ABSOLUTE';
        AxisData.Diag.sWaitReason := 'Waiting MC_MoveAbsolute.Done';
        AxisData.Diag.tStepPreset := AxisData.Timeouts.tMoveTimeout;

        xPowerRequest := TRUE;
        xMoveAbsExecute := TRUE;

        IF NOT AxisData.Command.xPowerPermit THEN
            xMoveAbsExecute := FALSE;
            AxisData.Error.dwLogicalErrorLatched :=
                AxisData.Error.dwLogicalErrorLatched OR LOG_POWER_PERMIT_LOST;
            AxisData.Diag.iLastErrorStep := TO_INT(AxisData.Diag.iStep);
            AxisData.Diag.iStep := E_AXIS_STATE.STOPPING;

        ELSIF AxisData.Command.xGlobalError THEN
            xMoveAbsExecute := FALSE;
            AxisData.Error.dwLogicalErrorLatched :=
                AxisData.Error.dwLogicalErrorLatched OR LOG_GLOBAL_DURING_MOTION;
            AxisData.Diag.iLastErrorStep := TO_INT(AxisData.Diag.iStep);
            AxisData.Diag.iStep := E_AXIS_STATE.STOPPING;

        ELSIF rtStop.Q THEN
            xMoveAbsExecute := FALSE;
            AxisData.Diag.iStep := E_AXIS_STATE.STOPPING;

        ELSIF fbMoveAbsolute.Error THEN
            xMoveAbsExecute := FALSE;
            AxisData.Error.dwAxisErrorLatched :=
                AxisData.Error.dwAxisErrorLatched OR AXE_MC_MOVE_ABS_ERROR;
            AxisData.Diag.udiLastErrorID := TO_UDINT(fbMoveAbsolute.ErrorID);
            AxisData.Diag.iLastErrorStep := TO_INT(AxisData.Diag.iStep);
            AxisData.Diag.iStep := E_AXIS_STATE.ERROR_RESET_MANAGER;

        ELSIF fbMoveAbsolute.CommandAborted THEN
            xMoveAbsExecute := FALSE;
            AxisData.Error.dwAxisErrorLatched :=
                AxisData.Error.dwAxisErrorLatched OR AXE_COMMAND_ABORTED;
            AxisData.Diag.udiLastErrorID := 3003;
            AxisData.Diag.iLastErrorStep := TO_INT(AxisData.Diag.iStep);
            AxisData.Diag.iStep := E_AXIS_STATE.ERROR_RESET_MANAGER;

        ELSIF xAxisErrorActual THEN
            xMoveAbsExecute := FALSE;
            AxisData.Error.dwAxisErrorLatched :=
                AxisData.Error.dwAxisErrorLatched OR AxisData.Error.dwAxisErrorActual;
            AxisData.Diag.iLastErrorStep := TO_INT(AxisData.Diag.iStep);
            AxisData.Diag.iStep := E_AXIS_STATE.ERROR_RESET_MANAGER;

        ELSIF fbMoveAbsolute.Done THEN
            xMoveAbsExecute := FALSE;
            AxisData.Status.xDone := TRUE;
            AxisData.Diag.iStep := E_AXIS_STATE.READY;
        END_IF;

    // --------------------------------------------------
    E_AXIS_STATE.MOVE_RELATIVE:
    // --------------------------------------------------
        AxisData.Diag.sStepName := 'MOVING_RELATIVE';
        AxisData.Diag.sWaitReason := 'Waiting MC_MoveRelative.Done';
        AxisData.Diag.tStepPreset := AxisData.Timeouts.tMoveTimeout;

        xPowerRequest := TRUE;
        xMoveRelExecute := TRUE;

        IF NOT AxisData.Command.xPowerPermit THEN
            xMoveRelExecute := FALSE;
            AxisData.Error.dwLogicalErrorLatched :=
                AxisData.Error.dwLogicalErrorLatched OR LOG_POWER_PERMIT_LOST;
            AxisData.Diag.iLastErrorStep := TO_INT(AxisData.Diag.iStep);
            AxisData.Diag.iStep := E_AXIS_STATE.STOPPING;

        ELSIF AxisData.Command.xGlobalError THEN
            xMoveRelExecute := FALSE;
            AxisData.Error.dwLogicalErrorLatched :=
                AxisData.Error.dwLogicalErrorLatched OR LOG_GLOBAL_DURING_MOTION;
            AxisData.Diag.iLastErrorStep := TO_INT(AxisData.Diag.iStep);
            AxisData.Diag.iStep := E_AXIS_STATE.STOPPING;

        ELSIF rtStop.Q THEN
            xMoveRelExecute := FALSE;
            AxisData.Diag.iStep := E_AXIS_STATE.STOPPING;

        ELSIF fbMoveRelative.Error THEN
            xMoveRelExecute := FALSE;
            AxisData.Error.dwAxisErrorLatched :=
                AxisData.Error.dwAxisErrorLatched OR AXE_MC_MOVE_REL_ERROR;
            AxisData.Diag.udiLastErrorID := TO_UDINT(fbMoveRelative.ErrorID);
            AxisData.Diag.iLastErrorStep := TO_INT(AxisData.Diag.iStep);
            AxisData.Diag.iStep := E_AXIS_STATE.ERROR_RESET_MANAGER;

        ELSIF fbMoveRelative.CommandAborted THEN
            xMoveRelExecute := FALSE;
            AxisData.Error.dwAxisErrorLatched :=
                AxisData.Error.dwAxisErrorLatched OR AXE_COMMAND_ABORTED;
            AxisData.Diag.udiLastErrorID := 3003;
            AxisData.Diag.iLastErrorStep := TO_INT(AxisData.Diag.iStep);
            AxisData.Diag.iStep := E_AXIS_STATE.ERROR_RESET_MANAGER;

        ELSIF xAxisErrorActual THEN
            xMoveRelExecute := FALSE;
            AxisData.Error.dwAxisErrorLatched :=
                AxisData.Error.dwAxisErrorLatched OR AxisData.Error.dwAxisErrorActual;
            AxisData.Diag.iLastErrorStep := TO_INT(AxisData.Diag.iStep);
            AxisData.Diag.iStep := E_AXIS_STATE.ERROR_RESET_MANAGER;

        ELSIF fbMoveRelative.Done THEN
            xMoveRelExecute := FALSE;
            AxisData.Status.xDone := TRUE;
            AxisData.Diag.iStep := E_AXIS_STATE.READY;
        END_IF;

    // --------------------------------------------------
    E_AXIS_STATE.STOPPING:
    // --------------------------------------------------
        AxisData.Diag.sStepName := 'STOPPING';
        AxisData.Diag.sWaitReason := 'Waiting MC_Stop.Done';
        AxisData.Diag.tStepPreset := AxisData.Timeouts.tStopTimeout;

        xPowerRequest := TRUE;
        xStopExecute := TRUE;

        IF fbStop.Error THEN
            xStopExecute := FALSE;
            AxisData.Error.dwAxisErrorLatched :=
                AxisData.Error.dwAxisErrorLatched OR AXE_MC_STOP_ERROR;
            AxisData.Diag.udiLastErrorID := TO_UDINT(fbStop.ErrorID);
            AxisData.Diag.iLastErrorStep := TO_INT(AxisData.Diag.iStep);
            AxisData.Diag.iStep := E_AXIS_STATE.ERROR_RESET_MANAGER;

        ELSIF fbStop.Done THEN
            AxisData.Status.xDone := TRUE;
            AxisData.Diag.iStep := E_AXIS_STATE.STOP_RELEASE;
        END_IF;

    // --------------------------------------------------
    E_AXIS_STATE.STOP_RELEASE:
    // --------------------------------------------------
        AxisData.Diag.sStepName := 'STOP_RELEASE';
        AxisData.Diag.sWaitReason := 'Releasing MC_Stop.Execute';
        AxisData.Diag.tStepPreset := T#1S;

        xPowerRequest := TRUE;
        xStopExecute := FALSE;

        IF NOT fbStop.Busy THEN
            IF AxisData.Command.xGlobalError OR
               (AxisData.Error.dwAxisErrorLatched <> DWORD#0) OR
               (AxisData.Error.dwLogicalErrorLatched <> DWORD#0) OR
               xAxisErrorActual
            THEN
                AxisData.Diag.iStep := E_AXIS_STATE.ERROR_RESET_MANAGER;
            ELSE
                AxisData.Diag.iStep := E_AXIS_STATE.READY;
            END_IF;
        END_IF;

    // --------------------------------------------------
    E_AXIS_STATE.ERROR_RESET_MANAGER:
    // --------------------------------------------------
        AxisData.Diag.sStepName := 'ERROR';
        AxisData.Diag.tStepPreset := T#0S;

        xResetExecute    := FALSE;
        xStopExecute     := FALSE;
        xHomeExecute     := FALSE;
        xMoveAbsExecute  := FALSE;
        xMoveRelExecute  := FALSE;
        xJogForwardExec  := FALSE;
        xJogBackwardExec := FALSE;

        IF AxisData.Timeouts.xDisableOnError THEN
            xPowerRequest := FALSE;
        ELSE
            xPowerRequest := AxisData.Command.xPowerPermit AND NOT xAxisErrorActual;
        END_IF;

        IF (AxisData.Error.dwAxisError = DWORD#0) AND
           (AxisData.Error.dwLogicalError = DWORD#0) AND
           NOT AxisData.Command.xGlobalError
        THEN
            AxisData.Diag.iStep := E_AXIS_STATE.DISABLED;

        ELSE
            IF AxisData.Command.xGlobalError THEN
                AxisData.Diag.sWaitReason := 'Waiting global error release';
            ELSIF (AxisData.Error.dwAxisError <> DWORD#0) AND
                  (AxisData.Error.dwLogicalError <> DWORD#0) THEN
                AxisData.Diag.sWaitReason := 'Waiting ResetAllError';
            ELSIF AxisData.Error.dwAxisError <> DWORD#0 THEN
                AxisData.Diag.sWaitReason := 'Waiting ResetAxisError or ResetAllError';
            ELSIF AxisData.Error.dwLogicalError <> DWORD#0 THEN
                AxisData.Diag.sWaitReason := 'Waiting ResetLogicalError or ResetAllError';
            ELSE
                AxisData.Diag.sWaitReason := 'Waiting reset';
            END_IF;

            IF rtResetAllError.Q AND xResetPermit THEN
                xDoResetAxis := TRUE;
                xDoResetLogical := TRUE;
                IF xNeedMcReset THEN
                    AxisData.Diag.iStep := E_AXIS_STATE.RESET_AXIS_ERROR;
                ELSE
                    AxisData.Diag.iStep := E_AXIS_STATE.RESET_FINISH;
                END_IF;

            ELSIF rtResetAxisError.Q THEN
                xDoResetAxis := TRUE;
                xDoResetLogical := FALSE;
                IF xNeedMcReset THEN
                    AxisData.Diag.iStep := E_AXIS_STATE.RESET_AXIS_ERROR;
                ELSE
                    AxisData.Diag.iStep := E_AXIS_STATE.RESET_FINISH;
                END_IF;

            ELSIF rtResetLogicalError.Q THEN
                xDoResetAxis := FALSE;
                xDoResetLogical := TRUE;
                AxisData.Diag.iStep := E_AXIS_STATE.RESET_FINISH;
            END_IF;
        END_IF;

    // --------------------------------------------------
    E_AXIS_STATE.RESET_AXIS_ERROR:
    // --------------------------------------------------
        AxisData.Diag.sStepName := 'RESET_AXIS_ERROR';
        AxisData.Diag.sWaitReason := 'Waiting MC_Reset.Done';
        AxisData.Diag.tStepPreset := AxisData.Timeouts.tResetTimeout;

        xPowerRequest := FALSE;
        xResetExecute := TRUE;

        IF fbReset.Error THEN
            AxisData.Diag.sWarningText := 'MC_Reset finished with error';
            uiResetWarningCode := WRN_RESET_MC_ERROR;
            xResetExecute := FALSE;
            AxisData.Error.dwAxisErrorLatched :=
                AxisData.Error.dwAxisErrorLatched OR AXE_MC_RESET_ERROR;
            AxisData.Diag.udiLastErrorID := TO_UDINT(fbReset.ErrorID);
            AxisData.Diag.iLastErrorStep := TO_INT(AxisData.Diag.iStep);
            AxisData.Diag.iStep := E_AXIS_STATE.ERROR_RESET_MANAGER;

        ELSIF fbReset.Done THEN
            xResetExecute := FALSE;
            AxisData.Diag.iStep := E_AXIS_STATE.RESET_RELEASE;
        END_IF;

    // --------------------------------------------------
    E_AXIS_STATE.RESET_RELEASE:
    // --------------------------------------------------
        AxisData.Diag.sStepName := 'RESET_RELEASE';
        AxisData.Diag.sWaitReason := 'Releasing MC_Reset.Execute';
        AxisData.Diag.tStepPreset := T#1S;

        xPowerRequest := FALSE;
        xResetExecute := FALSE;

        IF NOT fbReset.Busy THEN
            AxisData.Diag.iStep := E_AXIS_STATE.RESET_FINISH;
        END_IF;

    // --------------------------------------------------
    E_AXIS_STATE.RESET_FINISH:
    // --------------------------------------------------
        AxisData.Diag.sStepName := 'RESET_FINISH';
        AxisData.Diag.sWaitReason := 'Finishing reset';
        AxisData.Diag.tStepPreset := T#0S;

        xPowerRequest := FALSE;
        xResetExecute := FALSE;

        IF xDoResetAxis THEN
            AxisData.Error.dwAxisErrorLatched := DWORD#0;
        END_IF;
        IF xDoResetLogical THEN
            AxisData.Error.dwLogicalErrorLatched := DWORD#0;
            AxisData.Diag.xStepTimeout := FALSE;
        END_IF;

        xDoResetAxis := FALSE;
        xDoResetLogical := FALSE;

        // Финальная проверка
        IF AxisData.Error.dwAxisErrorActual <> DWORD#0 THEN
            AxisData.Diag.sWarningText := 'Axis error remains active after reset';
            uiResetWarningCode := WRN_RESET_AXIS_ACTIVE;
            AxisData.Error.dwAxisErrorLatched :=
                AxisData.Error.dwAxisErrorLatched OR AxisData.Error.dwAxisErrorActual;
            AxisData.Diag.iStep := E_AXIS_STATE.ERROR_RESET_MANAGER;

        ELSIF AxisData.Error.dwAxisErrorLatched <> DWORD#0 THEN
            AxisData.Diag.sWarningText := 'Latched axis error was not reset';
            uiResetWarningCode := WRN_RESET_AXIS_LATCHED;
            AxisData.Diag.iStep := E_AXIS_STATE.ERROR_RESET_MANAGER;

        ELSIF AxisData.Error.dwLogicalErrorLatched <> DWORD#0 THEN
            AxisData.Diag.sWarningText := 'Logical axis error was not reset';
            uiResetWarningCode := WRN_RESET_LOGICAL_ACTIVE;
            AxisData.Diag.iStep := E_AXIS_STATE.ERROR_RESET_MANAGER;

        ELSIF AxisData.Command.xGlobalError THEN
            AxisData.Diag.sWarningText := 'Global error is still active';
            uiResetWarningCode := WRN_RESET_GLOBAL_ERROR;
            AxisData.Diag.iStep := E_AXIS_STATE.ERROR_RESET_MANAGER;

        ELSE
            AxisData.Diag.iStep := E_AXIS_STATE.DISABLED;
        END_IF;

    // --------------------------------------------------
    ELSE  // неизвестное состояние
    // --------------------------------------------------
        AxisData.Error.dwLogicalErrorLatched :=
            AxisData.Error.dwLogicalErrorLatched OR LOG_UNKNOWN_STEP;
        AxisData.Diag.iLastErrorStep := TO_INT(AxisData.Diag.iStep);
        AxisData.Diag.iStep := E_AXIS_STATE.ERROR_RESET_MANAGER;

END_CASE;

// ======================================================
// 5. ТАЙМЕР ШАГА И КОНТРОЛЬ ТАЙМАУТА
// ======================================================
xStepChanged := (AxisData.Diag.iStep <> iPrevStep);
IF xStepChanged THEN
    iPrevStep := AxisData.Diag.iStep;
    xStepTimerEnable := FALSE;
ELSE
    xStepTimerEnable := TRUE;
END_IF;

tonStep(IN := xStepTimerEnable, PT := T#1000H);
AxisData.Diag.tStepElapsed := tonStep.ET;

tonStepTimeout(
    IN := xStepTimerEnable AND (AxisData.Diag.tStepPreset > T#0S),
    PT := AxisData.Diag.tStepPreset
);

IF tonStepTimeout.Q AND (AxisData.Diag.iStep <> E_AXIS_STATE.ERROR_RESET_MANAGER) THEN
    IF (AxisData.Diag.iStep = E_AXIS_STATE.RESET_AXIS_ERROR)
    OR (AxisData.Diag.iStep = E_AXIS_STATE.RESET_RELEASE) THEN
        AxisData.Diag.sWarningText := 'Axis reset timeout';
        uiResetWarningCode := WRN_RESET_TIMEOUT;
    END_IF;

    AxisData.Diag.xStepTimeout := TRUE;
    AxisData.Error.dwLogicalErrorLatched := AxisData.Error.dwLogicalErrorLatched OR LOG_STEP_TIMEOUT;
    AxisData.Diag.iLastErrorStep := TO_INT(AxisData.Diag.iStep);

    xResetExecute    := FALSE;
    xStopExecute     := FALSE;
    xHomeExecute     := FALSE;
    xMoveAbsExecute  := FALSE;
    xMoveRelExecute  := FALSE;
    xJogForwardExec  := FALSE;
    xJogBackwardExec := FALSE;

    AxisData.Diag.iStep := E_AXIS_STATE.ERROR_RESET_MANAGER;
END_IF;

IF uiResetWarningCode <> UINT#0 THEN
    AxisData.Diag.stWarning.uiCode := uiResetWarningCode;
    AxisData.Diag.stWarning.udiSequence := AxisData.Diag.stWarning.udiSequence + UDINT#1;
    IF AxisData.Diag.stWarning.udiSequence = UDINT#0 THEN
        AxisData.Diag.stWarning.udiSequence := UDINT#1;
    END_IF;
    xWarningPulse := TRUE;
END_IF;

// ======================================================
// 6. УДЕРЖАНИЕ ПРЕДУПРЕЖДЕНИЙ (TP)
// ======================================================
tpWarningHold(IN := xWarningPulse, PT := T#2S);
IF NOT tpWarningHold.Q THEN
    AxisData.Error.dwWarningLatched := DWORD#0;
    AxisData.Diag.sWarningText := '';
END_IF;
AxisData.Error.dwWarning := AxisData.Error.dwWarningLatched;
AxisData.Status.xWarning := (AxisData.Error.dwWarning <> DWORD#0);

// ======================================================
// 7. ВЫЗОВ MC-БЛОКОВ
// ======================================================
fbPower(
    Axis := Axis,
    // Enable активирует обработку MC_Power и не является командой питания.
    // Для штатного выключения FB продолжает выполняться, а силовые входы снимаются.
    Enable := TRUE,
    bRegulatorOn := xPowerRequest,
    bDriveStart := xPowerRequest
);

fbReset(
    Axis := Axis,
    Execute := xResetExecute
);

fbStop(
    Axis := Axis,
    Execute := xStopExecute,
    Deceleration := lrEffectiveDeceleration,
    Jerk := lrEffectiveJerk
);

fbJog(
    Axis := Axis,
    JogForward := xJogForwardExec,
    JogBackward := xJogBackwardExec,
    Velocity := lrEffectiveVelocity,
    Acceleration := lrEffectiveAcceleration,
    Deceleration := lrEffectiveDeceleration,
    Jerk := lrEffectiveJerk
);

fbHome(
    Axis := Axis,
    Execute := xHomeExecute,
    Position := AxisData.MotionParam.lrHomePosition
);

fbMoveAbsolute(
    Axis := Axis,
    Execute := xMoveAbsExecute,
    Position := AxisData.MotionParam.lrTargetPosition,
    Velocity := lrEffectiveVelocity,
    Acceleration := lrEffectiveAcceleration,
    Deceleration := lrEffectiveDeceleration,
    Jerk := lrEffectiveJerk,
    Direction := MC_DIRECTION.shortest,
    BufferMode := MC_BUFFER_MODE.Aborting
);

fbMoveRelative(
    Axis := Axis,
    Execute := xMoveRelExecute,
    Distance := AxisData.MotionParam.lrDistance,
    Velocity := lrEffectiveVelocity,
    Acceleration := lrEffectiveAcceleration,
    Deceleration := lrEffectiveDeceleration,
    Jerk := lrEffectiveJerk,
    BufferMode := MC_BUFFER_MODE.Aborting
);

fbReadPosition(
    Axis := Axis,
    Enable := TRUE
);

fbReadStatus(
    Axis := Axis,
    Enable := TRUE
);

fbReadAxisError(
    Axis := Axis,
    Enable := TRUE
);

// ======================================================
// 8. ИТОГОВЫЕ СТАТУСЫ (запись в структуру)
// ======================================================
AxisData.Status.xStandstill := fbReadStatus.Valid AND NOT AxisData.Status.xMotionBusy
	AND (fbReadStatus.StandStill OR fbReadStatus.Disabled OR fbReadStatus.Errorstop);
AxisData.Status.lrActualPosition := LREAL_TO_REAL(fbReadPosition.Position);

// Повторно собираем актуальные ошибки (для полноты)
AxisData.Error.dwAxisErrorActual := DWORD#0;
AxisData.Error.dwAxisErrorActual.0  := fbPower.Error;
AxisData.Error.dwAxisErrorActual.1  := fbReset.Error;
AxisData.Error.dwAxisErrorActual.2  := fbStop.Error;
AxisData.Error.dwAxisErrorActual.3  := fbJog.Error;
AxisData.Error.dwAxisErrorActual.4  := fbHome.Error;
AxisData.Error.dwAxisErrorActual.5  := fbMoveAbsolute.Error;
AxisData.Error.dwAxisErrorActual.6  := fbMoveRelative.Error;
AxisData.Error.dwAxisErrorActual.7  := fbReadPosition.Error;
AxisData.Error.dwAxisErrorActual.8  := fbReadStatus.Error;
AxisData.Error.dwAxisErrorActual.9  := fbReadStatus.Errorstop;
AxisData.Error.dwAxisErrorActual.10 := fbReadStatus.FBErrorOccured;
AxisData.Error.dwAxisErrorActual.11 := fbReadAxisError.AxisError;

xAxisErrorActual := (AxisData.Error.dwAxisErrorActual <> DWORD#0);

AxisData.Status.xLocalError :=
    fbPower.Error OR
    fbReset.Error OR
    fbStop.Error OR
    fbJog.Error OR
    fbHome.Error OR
    fbMoveAbsolute.Error OR
    fbMoveRelative.Error OR
    fbReadPosition.Error OR
    fbReadStatus.Error OR
    fbReadStatus.Errorstop OR
    fbReadStatus.FBErrorOccured OR
    fbReadAxisError.AxisError;

AxisData.Status.xMotionBusy :=
    fbStop.Busy OR
    fbJog.Busy OR
    fbHome.Busy OR
    fbMoveAbsolute.Busy OR
    fbMoveRelative.Busy;

xNeedMcReset :=
    fbReadStatus.Errorstop OR
    fbReadStatus.FBErrorOccured OR
    fbReadAxisError.AxisError;

AxisData.Error.dwAxisError := AxisData.Error.dwAxisErrorActual OR AxisData.Error.dwAxisErrorLatched;
AxisData.Error.dwLogicalError := AxisData.Error.dwLogicalErrorLatched;
AxisData.Error.dwAllError := AxisData.Error.dwAxisError OR AxisData.Error.dwLogicalError;
AxisData.Error.dwAlarmActive := AxisData.Error.dwAxisError
    OR SHL(AxisData.Error.dwLogicalError, 16);
AxisData.Error.dwDriveAxisErrorID := fbReadAxisError.AxisErrorID;

AxisData.Status.xAxisError := (AxisData.Error.dwAxisError <> DWORD#0);
AxisData.Status.xLogicalError := (AxisData.Error.dwLogicalError <> DWORD#0);
AxisData.Status.xAxisResetNeeded := AxisData.Status.xAxisError;
AxisData.Status.xLogicalResetNeeded := AxisData.Status.xLogicalError;

AxisData.Status.xError :=
    (AxisData.Diag.iStep = E_AXIS_STATE.ERROR_RESET_MANAGER) OR
    AxisData.Status.xAxisError OR
    AxisData.Status.xLogicalError OR
    AxisData.Command.xGlobalError;

AxisData.Status.xBusy :=
    fbPower.Busy OR
    fbReset.Busy OR
    AxisData.Status.xMotionBusy;

AxisData.Status.xCanStartMotion :=
    (AxisData.Diag.iStep = E_AXIS_STATE.READY) AND
    AxisData.Status.xPowered AND
    NOT AxisData.Status.xMotionBusy AND
    NOT AxisData.Status.xAxisError AND
    NOT AxisData.Status.xLogicalError AND
    NOT AxisData.Command.xGlobalError;

// ======================================================
// 9. ТЕКСТ ОШИБКИ И ID
// ======================================================
AxisData.Diag.sErrorText := '';
AxisData.Diag.udiActualErrorID := 0;

IF (AxisData.Error.dwLogicalError AND LOG_POWER_PERMIT_LOST) <> DWORD#0 THEN
    AxisData.Diag.sErrorText := 'Power permit lost';
    AxisData.Diag.udiActualErrorID := 1001;

ELSIF (AxisData.Error.dwLogicalError AND LOG_GLOBAL_DURING_POWER) <> DWORD#0 THEN
    AxisData.Diag.sErrorText := 'Global error during power on';
    AxisData.Diag.udiActualErrorID := 1002;

ELSIF (AxisData.Error.dwLogicalError AND LOG_GLOBAL_DURING_READY) <> DWORD#0 THEN
    AxisData.Diag.sErrorText := 'Global error in READY state';
    AxisData.Diag.udiActualErrorID := 2000;

ELSIF (AxisData.Error.dwLogicalError AND LOG_GLOBAL_DURING_MOTION) <> DWORD#0 THEN
    AxisData.Diag.sErrorText := 'Global error during motion';
    AxisData.Diag.udiActualErrorID := 2100;

ELSIF (AxisData.Error.dwLogicalError AND LOG_JOG_CONFLICT) <> DWORD#0 THEN
    AxisData.Diag.sErrorText := 'Jog positive and negative active together';
    AxisData.Diag.udiActualErrorID := 2001;

ELSIF (AxisData.Error.dwLogicalError AND LOG_MOVE_ABS_NOT_HOMED) <> DWORD#0 THEN
    AxisData.Diag.sErrorText := 'MoveAbsolute denied: axis not homed';
    AxisData.Diag.udiActualErrorID := 1200;

ELSIF (AxisData.Error.dwLogicalError AND LOG_MOVE_REL_NOT_HOMED) <> DWORD#0 THEN
    AxisData.Diag.sErrorText := 'MoveRelative denied: axis not homed';
    AxisData.Diag.udiActualErrorID := 1300;

ELSIF (AxisData.Error.dwLogicalError AND LOG_STEP_TIMEOUT) <> DWORD#0 THEN
    AxisData.Diag.sErrorText := 'Step timeout';
    AxisData.Diag.udiActualErrorID := 9000 + INT_TO_UDINT(AxisData.Diag.iLastErrorStep);

ELSIF (AxisData.Error.dwLogicalError AND LOG_UNKNOWN_STEP) <> DWORD#0 THEN
    AxisData.Diag.sErrorText := 'Unknown axis step';
    AxisData.Diag.udiActualErrorID := 9999;

ELSIF (AxisData.Error.dwAxisError AND AXE_MC_POWER_ERROR) <> DWORD#0 THEN
    AxisData.Diag.sErrorText := 'MC_Power error';
    AxisData.Diag.udiActualErrorID := TO_UDINT(fbPower.ErrorID);

ELSIF (AxisData.Error.dwAxisError AND AXE_MC_RESET_ERROR) <> DWORD#0 THEN
    AxisData.Diag.sErrorText := 'MC_Reset error';
    AxisData.Diag.udiActualErrorID := TO_UDINT(fbReset.ErrorID);

ELSIF (AxisData.Error.dwAxisError AND AXE_MC_STOP_ERROR) <> DWORD#0 THEN
    AxisData.Diag.sErrorText := 'MC_Stop error';
    AxisData.Diag.udiActualErrorID := TO_UDINT(fbStop.ErrorID);

ELSIF (AxisData.Error.dwAxisError AND AXE_MC_JOG_ERROR) <> DWORD#0 THEN
    AxisData.Diag.sErrorText := 'MC_Jog error';
    AxisData.Diag.udiActualErrorID := TO_UDINT(fbJog.ErrorID);

ELSIF (AxisData.Error.dwAxisError AND AXE_MC_HOME_ERROR) <> DWORD#0 THEN
    AxisData.Diag.sErrorText := 'MC_Home error';
    AxisData.Diag.udiActualErrorID := TO_UDINT(fbHome.ErrorID);

ELSIF (AxisData.Error.dwAxisError AND AXE_MC_MOVE_ABS_ERROR) <> DWORD#0 THEN
    AxisData.Diag.sErrorText := 'MC_MoveAbsolute error';
    AxisData.Diag.udiActualErrorID := TO_UDINT(fbMoveAbsolute.ErrorID);

ELSIF (AxisData.Error.dwAxisError AND AXE_MC_MOVE_REL_ERROR) <> DWORD#0 THEN
    AxisData.Diag.sErrorText := 'MC_MoveRelative error';
    AxisData.Diag.udiActualErrorID := TO_UDINT(fbMoveRelative.ErrorID);

ELSIF (AxisData.Error.dwAxisError AND AXE_READ_POS_ERROR) <> DWORD#0 THEN
    AxisData.Diag.sErrorText := 'MC_ReadActualPosition error';
    AxisData.Diag.udiActualErrorID := TO_UDINT(fbReadPosition.ErrorID);

ELSIF (AxisData.Error.dwAxisError AND AXE_READ_STATUS_ERROR) <> DWORD#0 THEN
    AxisData.Diag.sErrorText := 'MC_ReadStatus error';
    AxisData.Diag.udiActualErrorID := TO_UDINT(fbReadStatus.ErrorID);

ELSIF (AxisData.Error.dwAxisError AND AXE_ERRORSTOP) <> DWORD#0 THEN
    AxisData.Diag.sErrorText := 'Axis Errorstop active';
    AxisData.Diag.udiActualErrorID := 3001;

ELSIF (AxisData.Error.dwAxisError AND AXE_FB_ERROR_OCCURRED) <> DWORD#0 THEN
    AxisData.Diag.sErrorText := 'SoftMotion FBErrorOccured active';
    AxisData.Diag.udiActualErrorID := 3002;

ELSIF (AxisData.Error.dwAxisError AND AXE_COMMAND_ABORTED) <> DWORD#0 THEN
    AxisData.Diag.sErrorText := 'Motion command aborted';
    AxisData.Diag.udiActualErrorID := 3003;

ELSIF (AxisData.Error.dwAxisError AND AXE_UNKNOWN_ACTUAL_ERROR) <> DWORD#0 THEN
    AxisData.Diag.sErrorText := 'Unknown actual axis error';
    AxisData.Diag.udiActualErrorID := 3004;

ELSIF (AxisData.Error.dwAxisError AND AXE_DRIVE_AXIS_ERROR) <> DWORD#0 THEN
    AxisData.Diag.sErrorText := 'Drive axis error active';
    AxisData.Diag.udiActualErrorID := DWORD_TO_UDINT(fbReadAxisError.AxisErrorID);

ELSIF (AxisData.Error.dwAxisError AND AXE_POWER_FEEDBACK_LOST) <> DWORD#0 THEN
    AxisData.Diag.sErrorText := 'Drive power feedback lost';
    AxisData.Diag.udiActualErrorID := 3005;

ELSIF AxisData.Command.xGlobalError THEN
    AxisData.Diag.sErrorText := 'Global error active';
    AxisData.Diag.udiActualErrorID := 5000;
END_IF;

IF AxisData.Diag.udiActualErrorID <> 0 THEN
    AxisData.Diag.udiLastErrorID := AxisData.Diag.udiActualErrorID;
END_IF;

// Сохраняем последнюю ненулевую ошибку и формируем удобное представление для HMI.
IF (AxisData.Error.dwAxisError <> DWORD#0)
OR (AxisData.Error.dwLogicalError <> DWORD#0) THEN
	AxisData.Error.dwAxisErrorLast := AxisData.Error.dwAxisError;
	AxisData.Error.dwLogicalErrorLast := AxisData.Error.dwLogicalError;
END_IF;

AxisData.Error.stErrorActive := UpdateErrorView(
	dwAxisError := AxisData.Error.dwAxisError,
	dwLogicalError := AxisData.Error.dwLogicalError
);
AxisData.Error.stErrorLast := UpdateErrorView(
    dwAxisError := AxisData.Error.dwAxisErrorLast,
    dwLogicalError := AxisData.Error.dwLogicalErrorLast
);

FaultStatus.xResetAllowed := AxisData.Status.xError
	AND xResetPermit
	AND NOT AxisData.Command.xGlobalError
	AND NOT FaultStatus.xBusy;
